(* IEC 61131-3 sources: trust-platform/examples/OSCAT/refinery_temperature_conditioning/oop/src, 3 files *)

(* ---- Main.st ---- *)
(* Pattern role: ISignalSource is the contract boundary for the Decorator example. *)
INTERFACE ISignalSource EXTENDS IComponent
    PROPERTY Value : REAL
    GET
    END_GET
    END_PROPERTY

    PROPERTY Quality : BYTE
    GET
    END_GET
    END_PROPERTY

    METHOD Update
    END_METHOD
END_INTERFACE

(* Pattern role: RawAnalogInput is a concrete implementation in the Decorator example. *)
FUNCTION_BLOCK RawAnalogInput IMPLEMENTS ISignalSource
VAR
    ValueValue : REAL;
    QualityValue : BYTE;
    ReadyValue : BOOL;
    ErrorValue : BOOL;
    ErrorIdValue : WORD;
    StatusValue : BYTE;
END_VAR

METHOD PUBLIC Configure
VAR_INPUT
    InputValue : REAL;
    InputQuality : BYTE;
END_VAR
ValueValue := InputValue;
QualityValue := InputQuality;
END_METHOD

METHOD PUBLIC Initialize
ReadyValue := TRUE;
QualityValue := BYTE#2;
ClearError();
END_METHOD

METHOD PUBLIC Reset
ValueValue := REAL#0.0;
QualityValue := BYTE#2;
ClearError();
END_METHOD

METHOD PUBLIC ClearError
ErrorValue := FALSE;
ErrorIdValue := WORD#0;
StatusValue := BYTE#0;
END_METHOD

METHOD PUBLIC Snapshot : ComponentStatus
VAR
    Result : ComponentStatus;
END_VAR
Result.Ready := ReadyValue;
Result.Error := ErrorValue;
Result.ErrorId := ErrorIdValue;
Result.Status := StatusValue;
Snapshot := Result;
END_METHOD

METHOD PUBLIC Update
END_METHOD

PUBLIC PROPERTY Value : REAL
GET
    Value := ValueValue;
END_GET
END_PROPERTY

PUBLIC PROPERTY Quality : BYTE
GET
    Quality := QualityValue;
END_GET
END_PROPERTY

PUBLIC PROPERTY Ready : BOOL
GET
    Ready := ReadyValue;
END_GET
END_PROPERTY

PUBLIC PROPERTY Error : BOOL
GET
    Error := ErrorValue;
END_GET
END_PROPERTY

PUBLIC PROPERTY ErrorId : WORD
GET
    ErrorId := ErrorIdValue;
END_GET
END_PROPERTY

PUBLIC PROPERTY Status : BYTE
GET
    Status := StatusValue;
END_GET
END_PROPERTY
END_FUNCTION_BLOCK

(* Pattern role: VotingDecorator is a concrete implementation in the Decorator example. *)
FUNCTION_BLOCK VotingDecorator IMPLEMENTS ISignalSource
VAR
    Source1 : ISignalSource;
    Source2 : ISignalSource;
    Source3 : ISignalSource;
    ValueValue : REAL;
    QualityValue : BYTE;
    ReadyValue : BOOL;
    ErrorValue : BOOL;
    ErrorIdValue : WORD;
    StatusValue : BYTE;
END_VAR

METHOD PUBLIC SetSources
VAR_INPUT
    First : ISignalSource;
    Second : ISignalSource;
    Third : ISignalSource;
END_VAR
Source1 := First;
Source2 := Second;
Source3 := Third;
END_METHOD

METHOD PUBLIC Initialize
ReadyValue := TRUE;
QualityValue := BYTE#0;
ClearError();
END_METHOD

METHOD PUBLIC Reset
ValueValue := REAL#0.0;
QualityValue := BYTE#0;
ClearError();
END_METHOD

METHOD PUBLIC ClearError
ErrorValue := FALSE;
ErrorIdValue := WORD#0;
StatusValue := BYTE#0;
END_METHOD

METHOD PUBLIC Snapshot : ComponentStatus
VAR
    Result : ComponentStatus;
END_VAR
Result.Ready := ReadyValue;
Result.Error := ErrorValue;
Result.ErrorId := ErrorIdValue;
Result.Status := StatusValue;
Snapshot := Result;
END_METHOD

METHOD PUBLIC Update
Source1.Update();
Source2.Update();
Source3.Update();
IF (Source1.Quality = BYTE#2) AND (Source2.Quality = BYTE#2) THEN
    ValueValue := (Source1.Value + Source2.Value) / REAL#2.0;
    QualityValue := BYTE#2;
ELSIF (Source1.Quality = BYTE#2) AND (Source3.Quality = BYTE#2) THEN
    ValueValue := (Source1.Value + Source3.Value) / REAL#2.0;
    QualityValue := BYTE#2;
ELSIF (Source2.Quality = BYTE#2) AND (Source3.Quality = BYTE#2) THEN
    ValueValue := (Source2.Value + Source3.Value) / REAL#2.0;
    QualityValue := BYTE#2;
ELSE
    QualityValue := BYTE#0;
END_IF;
END_METHOD

PUBLIC PROPERTY Value : REAL
GET
    Value := ValueValue;
END_GET
END_PROPERTY

PUBLIC PROPERTY Quality : BYTE
GET
    Quality := QualityValue;
END_GET
END_PROPERTY

PUBLIC PROPERTY Ready : BOOL
GET
    Ready := ReadyValue;
END_GET
END_PROPERTY

PUBLIC PROPERTY Error : BOOL
GET
    Error := ErrorValue;
END_GET
END_PROPERTY

PUBLIC PROPERTY ErrorId : WORD
GET
    ErrorId := ErrorIdValue;
END_GET
END_PROPERTY

PUBLIC PROPERTY Status : BYTE
GET
    Status := StatusValue;
END_GET
END_PROPERTY
END_FUNCTION_BLOCK

(* Pattern role: RangeClampDecorator is a concrete implementation in the Decorator example. *)
FUNCTION_BLOCK RangeClampDecorator IMPLEMENTS ISignalSource
VAR
    Inner : ISignalSource;
    MinValue : REAL;
    MaxValue : REAL;
    ValueValue : REAL;
    QualityValue : BYTE;
    ClampFaultValue : BOOL;
    ReadyValue : BOOL;
    ErrorValue : BOOL;
    ErrorIdValue : WORD;
    StatusValue : BYTE;
END_VAR

METHOD PUBLIC Wrap
VAR_INPUT
    InnerSource : ISignalSource;
    Minimum : REAL;
    Maximum : REAL;
END_VAR
Inner := InnerSource;
MinValue := Minimum;
MaxValue := Maximum;
END_METHOD

METHOD PUBLIC Initialize
ReadyValue := TRUE;
ClearError();
END_METHOD

METHOD PUBLIC Reset
ValueValue := REAL#0.0;
QualityValue := BYTE#0;
ClampFaultValue := FALSE;
ClearError();
END_METHOD

METHOD PUBLIC ClearError
ErrorValue := FALSE;
ErrorIdValue := WORD#0;
StatusValue := BYTE#0;
END_METHOD

METHOD PUBLIC Snapshot : ComponentStatus
VAR
    Result : ComponentStatus;
END_VAR
Result.Ready := ReadyValue;
Result.Error := ErrorValue;
Result.ErrorId := ErrorIdValue;
Result.Status := StatusValue;
Snapshot := Result;
END_METHOD

METHOD PUBLIC Update
Inner.Update();
ClampFaultValue := FALSE;
IF Inner.Value < MinValue THEN
    ValueValue := MinValue;
    QualityValue := BYTE#0;
    ClampFaultValue := TRUE;
ELSIF Inner.Value > MaxValue THEN
    ValueValue := MaxValue;
    QualityValue := BYTE#0;
    ClampFaultValue := TRUE;
ELSE
    ValueValue := Inner.Value;
    QualityValue := Inner.Quality;
END_IF;
END_METHOD

PUBLIC PROPERTY ClampFault : BOOL
GET
    ClampFault := ClampFaultValue;
END_GET
END_PROPERTY

PUBLIC PROPERTY Value : REAL
GET
    Value := ValueValue;
END_GET
END_PROPERTY

PUBLIC PROPERTY Quality : BYTE
GET
    Quality := QualityValue;
END_GET
END_PROPERTY

PUBLIC PROPERTY Ready : BOOL
GET
    Ready := ReadyValue;
END_GET
END_PROPERTY

PUBLIC PROPERTY Error : BOOL
GET
    Error := ErrorValue;
END_GET
END_PROPERTY

PUBLIC PROPERTY ErrorId : WORD
GET
    ErrorId := ErrorIdValue;
END_GET
END_PROPERTY

PUBLIC PROPERTY Status : BYTE
GET
    Status := StatusValue;
END_GET
END_PROPERTY
END_FUNCTION_BLOCK

(* Pattern role: SpikeRejectDecorator is a concrete implementation in the Decorator example. *)
FUNCTION_BLOCK SpikeRejectDecorator IMPLEMENTS ISignalSource
VAR
    Inner : ISignalSource;
    MaxStepValue : REAL;
    ValueValue : REAL;
    QualityValue : BYTE;
    LastGoodValue : REAL;
    HasLastGood : BOOL;
    RejectedCountValue : INT;
    ReadyValue : BOOL;
    ErrorValue : BOOL;
    ErrorIdValue : WORD;
    StatusValue : BYTE;
END_VAR

METHOD PUBLIC Wrap
VAR_INPUT
    InnerSource : ISignalSource;
    MaxStep : REAL;
END_VAR
Inner := InnerSource;
MaxStepValue := MaxStep;
END_METHOD

METHOD PUBLIC Initialize
ReadyValue := TRUE;
ClearError();
END_METHOD

METHOD PUBLIC Reset
ValueValue := REAL#0.0;
QualityValue := BYTE#0;
LastGoodValue := REAL#0.0;
HasLastGood := FALSE;
RejectedCountValue := INT#0;
ClearError();
END_METHOD

METHOD PUBLIC ClearError
ErrorValue := FALSE;
ErrorIdValue := WORD#0;
StatusValue := BYTE#0;
END_METHOD

METHOD PUBLIC Snapshot : ComponentStatus
VAR
    Result : ComponentStatus;
END_VAR
Result.Ready := ReadyValue;
Result.Error := ErrorValue;
Result.ErrorId := ErrorIdValue;
Result.Status := StatusValue;
Snapshot := Result;
END_METHOD

METHOD PUBLIC Update
Inner.Update();
IF Inner.Quality <> BYTE#2 THEN
    ValueValue := Inner.Value;
    QualityValue := Inner.Quality;
ELSIF HasLastGood AND (ABS(Inner.Value - LastGoodValue) > MaxStepValue) THEN
    ValueValue := LastGoodValue;
    QualityValue := BYTE#1;
    RejectedCountValue := RejectedCountValue + INT#1;
ELSE
    ValueValue := Inner.Value;
    QualityValue := BYTE#2;
    LastGoodValue := Inner.Value;
    HasLastGood := TRUE;
END_IF;
END_METHOD

PUBLIC PROPERTY RejectedCount : INT
GET
    RejectedCount := RejectedCountValue;
END_GET
END_PROPERTY

PUBLIC PROPERTY Value : REAL
GET
    Value := ValueValue;
END_GET
END_PROPERTY

PUBLIC PROPERTY Quality : BYTE
GET
    Quality := QualityValue;
END_GET
END_PROPERTY

PUBLIC PROPERTY Ready : BOOL
GET
    Ready := ReadyValue;
END_GET
END_PROPERTY

PUBLIC PROPERTY Error : BOOL
GET
    Error := ErrorValue;
END_GET
END_PROPERTY

PUBLIC PROPERTY ErrorId : WORD
GET
    ErrorId := ErrorIdValue;
END_GET
END_PROPERTY

PUBLIC PROPERTY Status : BYTE
GET
    Status := StatusValue;
END_GET
END_PROPERTY
END_FUNCTION_BLOCK

(* Pattern role: Pt1SignalDecorator is a concrete implementation in the Decorator example. *)
FUNCTION_BLOCK Pt1SignalDecorator IMPLEMENTS ISignalSource
VAR
    Inner : ISignalSource;
    Filter : Pt1Filter;
    ValueValue : REAL;
    QualityValue : BYTE;
    ReadyValue : BOOL;
    ErrorValue : BOOL;
    ErrorIdValue : WORD;
    StatusValue : BYTE;
END_VAR

METHOD PUBLIC Wrap
VAR_INPUT
    InnerSource : ISignalSource;
    TimeConstant : TIME;
END_VAR
Inner := InnerSource;
Filter.Initialize();
Filter.Configure(TimeConstant := TimeConstant, Gain := REAL#1.0);
END_METHOD

METHOD PUBLIC Initialize
ReadyValue := TRUE;
Filter.Initialize();
ClearError();
END_METHOD

METHOD PUBLIC Reset
Filter.Reset();
ValueValue := REAL#0.0;
QualityValue := BYTE#0;
ClearError();
END_METHOD

METHOD PUBLIC ClearError
ErrorValue := FALSE;
ErrorIdValue := WORD#0;
StatusValue := BYTE#0;
END_METHOD

METHOD PUBLIC Snapshot : ComponentStatus
VAR
    Result : ComponentStatus;
END_VAR
Result.Ready := ReadyValue;
Result.Error := ErrorValue;
Result.ErrorId := ErrorIdValue;
Result.Status := StatusValue;
Snapshot := Result;
END_METHOD

METHOD PUBLIC Update
Inner.Update();
IF Inner.Quality = BYTE#2 THEN
    ValueValue := Filter.Update(Sample := Inner.Value);
    QualityValue := BYTE#2;
ELSE
    ValueValue := Inner.Value;
    QualityValue := Inner.Quality;
END_IF;
END_METHOD

PUBLIC PROPERTY Value : REAL
GET
    Value := ValueValue;
END_GET
END_PROPERTY

PUBLIC PROPERTY Quality : BYTE
GET
    Quality := QualityValue;
END_GET
END_PROPERTY

PUBLIC PROPERTY Ready : BOOL
GET
    Ready := ReadyValue;
END_GET
END_PROPERTY

PUBLIC PROPERTY Error : BOOL
GET
    Error := ErrorValue;
END_GET
END_PROPERTY

PUBLIC PROPERTY ErrorId : WORD
GET
    ErrorId := ErrorIdValue;
END_GET
END_PROPERTY

PUBLIC PROPERTY Status : BYTE
GET
    Status := StatusValue;
END_GET
END_PROPERTY
END_FUNCTION_BLOCK

(* Composition role: SignalConditioningPipeline owns the collaborating objects used by this Decorator example. *)
FUNCTION_BLOCK SignalConditioningPipeline
VAR
    Tc1 : RawAnalogInput;
    Tc2 : RawAnalogInput;
    Tc3 : RawAnalogInput;
    Voted : VotingDecorator;
    Clamped : RangeClampDecorator;
    SpikeRejected : SpikeRejectDecorator;
    Filtered : Pt1SignalDecorator;
    Conditioned : ISignalSource;
END_VAR

METHOD PUBLIC Initialize
Tc1.Initialize();
Tc2.Initialize();
Tc3.Initialize();
Voted.Initialize();
Clamped.Initialize();
SpikeRejected.Initialize();
Filtered.Initialize();
Voted.SetSources(First := Tc1, Second := Tc2, Third := Tc3);
Clamped.Wrap(InnerSource := Voted, Minimum := REAL#0.0, Maximum := REAL#400.0);
SpikeRejected.Wrap(InnerSource := Clamped, MaxStep := REAL#25.0);
Filtered.Wrap(InnerSource := SpikeRejected, TimeConstant := T#1s);
Conditioned := Filtered;
END_METHOD

METHOD PUBLIC Update : REAL
VAR_INPUT
    Input1 : REAL;
    Quality1 : BYTE;
    Input2 : REAL;
    Quality2 : BYTE;
    Input3 : REAL;
    Quality3 : BYTE;
END_VAR
Tc1.Configure(InputValue := Input1, InputQuality := Quality1);
Tc2.Configure(InputValue := Input2, InputQuality := Quality2);
Tc3.Configure(InputValue := Input3, InputQuality := Quality3);
Conditioned.Update();
Update := Conditioned.Value;
END_METHOD

PUBLIC PROPERTY ConditionedValue : REAL
GET
    ConditionedValue := Conditioned.Value;
END_GET
END_PROPERTY

PUBLIC PROPERTY Quality : BYTE
GET
    Quality := Conditioned.Quality;
END_GET
END_PROPERTY

PUBLIC PROPERTY RejectedCount : INT
GET
    RejectedCount := SpikeRejected.RejectedCount;
END_GET
END_PROPERTY

PUBLIC PROPERTY ClampFault : BOOL
GET
    ClampFault := Clamped.ClampFault;
END_GET
END_PROPERTY
END_FUNCTION_BLOCK

(* Scan role: Main wires the example objects and exposes the PLC call path under test. *)
PROGRAM Main
VAR
    Conditioning : SignalConditioningPipeline;
    Tc1Raw : INT;
    Tc2Raw : INT;
    Tc3Raw : INT;
    ConditionedRaw : INT;
    GoodQualityOut : BOOL;
END_VAR

Conditioning.Initialize();
ConditionedRaw := REAL_TO_INT(Conditioning.Update(Input1 := INT_TO_REAL(Tc1Raw), Quality1 := BYTE#2, Input2 := INT_TO_REAL(Tc2Raw), Quality2 := BYTE#2, Input3 := INT_TO_REAL(Tc3Raw), Quality3 := BYTE#2));
GoodQualityOut := Conditioning.Quality = BYTE#2;
END_PROGRAM

(* ---- Configuration.st ---- *)
CONFIGURATION RefineryTemperatureConditioningOopConfiguration
RESOURCE RefineryTemperatureConditioningOop ON PLC
    TASK MainTask (INTERVAL := T#100ms, PRIORITY := 1);
    PROGRAM Conditioning WITH MainTask : Main;
END_RESOURCE
VAR_CONFIG
    Conditioning.Tc1Raw AT %IW0 : INT;
    Conditioning.Tc2Raw AT %IW2 : INT;
    Conditioning.Tc3Raw AT %IW4 : INT;
    Conditioning.ConditionedRaw AT %QW0 : INT;
    Conditioning.GoodQualityOut AT %QX0.0 : BOOL;
END_VAR
END_CONFIGURATION

(* ---- Tests.st ---- *)
TEST_PROGRAM DecoratorPipelineRejectsSingleScanSpike
VAR
    Chain : SignalConditioningPipeline;
    Value : REAL;
END_VAR

Chain.Initialize();
Value := Chain.Update(Input1 := REAL#100.0, Quality1 := BYTE#2, Input2 := REAL#102.0, Quality2 := BYTE#2, Input3 := REAL#99.0, Quality3 := BYTE#2);
ASSERT_EQUAL(EXPECTED := BYTE#2, ACTUAL := Chain.Quality);
Value := Chain.Update(Input1 := REAL#180.0, Quality1 := BYTE#2, Input2 := REAL#181.0, Quality2 := BYTE#2, Input3 := REAL#182.0, Quality3 := BYTE#2);
ASSERT_EQUAL(EXPECTED := BYTE#1, ACTUAL := Chain.Quality);
ASSERT_EQUAL(EXPECTED := INT#1, ACTUAL := Chain.RejectedCount);
END_TEST_PROGRAM

TEST_PROGRAM DecoratorPipelineClampMarksBadQuality
VAR
    Chain : SignalConditioningPipeline;
    Value : REAL;
END_VAR

Chain.Initialize();
Value := Chain.Update(Input1 := REAL#450.0, Quality1 := BYTE#2, Input2 := REAL#452.0, Quality2 := BYTE#2, Input3 := REAL#451.0, Quality3 := BYTE#2);
ASSERT_EQUAL(EXPECTED := BYTE#0, ACTUAL := Chain.Quality);
ASSERT_TRUE(IN := Chain.ClampFault);
ASSERT_NEAR(EXPECTED := REAL#400.0, ACTUAL := Chain.ConditionedValue, DELTA := REAL#0.001);
END_TEST_PROGRAM

(* Pipeline recovery test: drives the same Chain through clamp/spike/
   recovered states. Catches bugs where decorator quality flags or
   rejected-spike counters fail to recover when the input returns to
   normal. *)
TEST_PROGRAM DecoratorPipelineRecoversAfterTransientFault
VAR
    Chain : SignalConditioningPipeline;
    Value : REAL;
    SpikeCount : INT;
END_VAR

Chain.Initialize();

(* Healthy reading - quality good *)
Value := Chain.Update(Input1 := REAL#100.0, Quality1 := BYTE#2, Input2 := REAL#102.0, Quality2 := BYTE#2, Input3 := REAL#99.0, Quality3 := BYTE#2);
ASSERT_EQUAL(EXPECTED := BYTE#2, ACTUAL := Chain.Quality);

(* Spike - quality drops, rejected count grows *)
Value := Chain.Update(Input1 := REAL#180.0, Quality1 := BYTE#2, Input2 := REAL#181.0, Quality2 := BYTE#2, Input3 := REAL#182.0, Quality3 := BYTE#2);
SpikeCount := Chain.RejectedCount;
ASSERT_TRUE(IN := SpikeCount >= INT#1);

(* Recovered reading near previous normal - quality must recover, not
   stay at degraded from the prior spike *)
Value := Chain.Update(Input1 := REAL#100.0, Quality1 := BYTE#2, Input2 := REAL#102.0, Quality2 := BYTE#2, Input3 := REAL#99.0, Quality3 := BYTE#2);
ASSERT_EQUAL(EXPECTED := BYTE#2, ACTUAL := Chain.Quality);
END_TEST_PROGRAM

(* Voting test: when one transmitter goes bad (Quality=0), the voted
   value is the average of the two good ones — not corrupted by the bad
   reading. The decorator chain still produces a good quality at the end. *)
TEST_PROGRAM DecoratorPipelineVotingTwoOfThree
VAR
    Chain : SignalConditioningPipeline;
    Value : REAL;
END_VAR

Chain.Initialize();
(* Tc2 is bad (quality 0 = bad), but Tc1 and Tc3 agree — pipeline must
   still produce good quality from the two-of-three vote. The bad Tc2
   raw value is wildly different but must not poison the voted result. *)
Value := Chain.Update(Input1 := REAL#100.0, Quality1 := BYTE#2, Input2 := REAL#9999.0, Quality2 := BYTE#0, Input3 := REAL#102.0, Quality3 := BYTE#2);
ASSERT_EQUAL(EXPECTED := BYTE#2, ACTUAL := Chain.Quality);
(* Voted value must be the average of Tc1 and Tc3 = 101.0, not influenced
   by Tc2's 9999. Filtered through PT1, but first sample passes through. *)
ASSERT_TRUE(IN := Chain.ConditionedValue < REAL#150.0);
ASSERT_TRUE(IN := Chain.ConditionedValue > REAL#50.0);
END_TEST_PROGRAM

(* Voting test: when two transmitters fail, the pipeline reports BAD
   quality and does not propagate any single good signal as if it were
   trustworthy. *)
TEST_PROGRAM DecoratorPipelineVotingFailsOnTwoBad
VAR
    Chain : SignalConditioningPipeline;
    Value : REAL;
END_VAR

Chain.Initialize();
(* Two of three thermocouples have bad quality — voting decorator
   cannot produce a good vote; pipeline must reflect bad quality. *)
Value := Chain.Update(Input1 := REAL#100.0, Quality1 := BYTE#2, Input2 := REAL#101.0, Quality2 := BYTE#0, Input3 := REAL#102.0, Quality3 := BYTE#0);
ASSERT_EQUAL(EXPECTED := BYTE#0, ACTUAL := Chain.Quality);
END_TEST_PROGRAM

(* Multi-cycle filtering: the PT1 stage settles toward the input over
   repeated cycles; verifies the inner filter state is preserved across
   Update calls (not reset by some decorator's Update side effect). *)
TEST_PROGRAM DecoratorPipelineFilterAccumulatesAcrossCycles
VAR
    Chain : SignalConditioningPipeline;
    Value : REAL;
    I : INT;
END_VAR

Chain.Initialize();
(* Establish a baseline at 100C *)
Value := Chain.Update(Input1 := REAL#100.0, Quality1 := BYTE#2, Input2 := REAL#100.0, Quality2 := BYTE#2, Input3 := REAL#100.0, Quality3 := BYTE#2);
(* Drive the input up to 110C and let the filter follow. After many
   identical samples the conditioned value must approach 110, never
   exceed it, and never drop back to the old baseline of 100. *)
FOR I := 1 TO 30 DO
    Value := Chain.Update(Input1 := REAL#110.0, Quality1 := BYTE#2, Input2 := REAL#110.0, Quality2 := BYTE#2, Input3 := REAL#110.0, Quality3 := BYTE#2);
END_FOR;
ASSERT_TRUE(IN := Chain.ConditionedValue >= REAL#100.0);
ASSERT_TRUE(IN := Chain.ConditionedValue <= REAL#110.0);
ASSERT_EQUAL(EXPECTED := BYTE#2, ACTUAL := Chain.Quality);
END_TEST_PROGRAM

(* Lower-bound clamp: negative readings must be clamped to 0 and marked
   bad quality (reading below physical range = sensor fault). *)
TEST_PROGRAM DecoratorPipelineLowerClampMarksBadQuality
VAR
    Chain : SignalConditioningPipeline;
    Value : REAL;
END_VAR

Chain.Initialize();
(* All three thermocouples report -10C — physically impossible for a
   distillation column overhead; clamp to 0, mark bad. *)
Value := Chain.Update(Input1 := REAL#-10.0, Quality1 := BYTE#2, Input2 := REAL#-10.0, Quality2 := BYTE#2, Input3 := REAL#-10.0, Quality3 := BYTE#2);
ASSERT_EQUAL(EXPECTED := BYTE#0, ACTUAL := Chain.Quality);
ASSERT_TRUE(IN := Chain.ClampFault);
ASSERT_NEAR(EXPECTED := REAL#0.0, ACTUAL := Chain.ConditionedValue, DELTA := REAL#0.001);
END_TEST_PROGRAM

(* Per-FB isolation: two pipelines running in parallel must not share
   filter state, last-good values, or rejected counts. *)
TEST_PROGRAM DecoratorPipelineParallelInstancesIndependent
VAR
    ChainA : SignalConditioningPipeline;
    ChainB : SignalConditioningPipeline;
    Value : REAL;
END_VAR

ChainA.Initialize();
ChainB.Initialize();
(* Drive ChainA into a spike-reject state *)
Value := ChainA.Update(Input1 := REAL#100.0, Quality1 := BYTE#2, Input2 := REAL#100.0, Quality2 := BYTE#2, Input3 := REAL#100.0, Quality3 := BYTE#2);
Value := ChainA.Update(Input1 := REAL#180.0, Quality1 := BYTE#2, Input2 := REAL#180.0, Quality2 := BYTE#2, Input3 := REAL#180.0, Quality3 := BYTE#2);
ASSERT_TRUE(IN := ChainA.RejectedCount >= INT#1);
(* ChainB stays steady - its rejected count must remain 0 *)
Value := ChainB.Update(Input1 := REAL#100.0, Quality1 := BYTE#2, Input2 := REAL#100.0, Quality2 := BYTE#2, Input3 := REAL#100.0, Quality3 := BYTE#2);
Value := ChainB.Update(Input1 := REAL#101.0, Quality1 := BYTE#2, Input2 := REAL#101.0, Quality2 := BYTE#2, Input3 := REAL#101.0, Quality3 := BYTE#2);
ASSERT_EQUAL(EXPECTED := INT#0, ACTUAL := ChainB.RejectedCount);
END_TEST_PROGRAM
